(* IEC 61131-3 sources: plc-iiot-stack/adapters/sd_mqtt_1_0/src/POUs/Adapters/FB_MqttClientSdMqtt, 14 files *)

(* ---- FB_MqttClientSdMqtt.decl.st ---- *)
// Назначение: адаптер I_MqttClient на библиотеку CODESYS-MQTT (github.com/stefandreyer/CODESYS-MQTT), релиз
//             «stable» (Project Information: MQTT 1.0.0.0, компания Stefan Dreyer, пространство имён SD_MQTT).
//             НЕ КОМПИЛИРОВАЛСЯ С РАБОЧЕЙ БИБЛИОТЕКОЙ: на CODESYS 3.5.17.30 у библиотеки нет зависимостей
//             (OSCAT BASIC 3.3.3.0, OSCAT NETWORK 1.30, «Common Helper for development» и системные
//             библиотеки точных версий 3.5.5–3.5.13), поэтому файл лежит вне src/ (docs/MANUAL_STEPS.md, раздел 9).
//             Сигнатуры взяты из объявлений библиотеки (HANDLE_MQTT, MQTTPublish, MQTTSubscribe, MQTT_IN_OUT).
//             Пул из PUB_POOL публикаторов: библиотека требует не менять топик и текст до done и пускает
//             публикацию по фронту send. Логин и пароль брокера версия 1.0.0.0 через входы не принимает —
//             Connect с непустым sUser отклоняется (MQTT_ERR_AUTH_UNSUPPORTED), а не подключается без пароля.
//             Завещание (LWT) версия строит сама из ClientID (WillTopicBase, ClientWillTopic, ClientWillMessage
//             до 30 символов): offline/lwt по data_schema 6 с ней не получить; флаг retain принятых сообщений
//             не виден (проверка retained шлюза команд не срабатывает).
// Автор:      kr0nsch
// Версия:     0.1.0
// Документ:   docs/plc_mqtt.md, раздел «Адаптер I_MqttClient»
FUNCTION_BLOCK FB_MqttClientSdMqtt IMPLEMENTS I_MqttClient
VAR_INPUT
    tTimeout : TIME := T#5S;                           // HANDLE_MQTT.TIMEOUT
END_VAR
VAR
    fbHandler : SD_MQTT.HANDLE_MQTT;
    stInOut : SD_MQTT.MQTT_IN_OUT;
    stInfo : SD_MQTT.MQTT_INFO;
    aPublishers : ARRAY[1..PUB_POOL] OF SD_MQTT.MQTTPublish;
    aPubTopic : ARRAY[1..PUB_POOL] OF STRING(GVL_Const.MQTT_TOPIC_LEN);
    aPubPayload : ARRAY[1..PUB_POOL] OF STRING(GVL_Const.MQTT_PAYLOAD_LEN);
    aPubLen : ARRAY[1..PUB_POOL] OF UDINT;
    aPubQos : ARRAY[1..PUB_POOL] OF SD_MQTT.QoS;
    aPubRetain : ARRAY[1..PUB_POOL] OF BOOL;
    aPubState : ARRAY[1..PUB_POOL] OF USINT;          // SLOT_FREE, SLOT_SENDING, SLOT_RELEASE
    fbSubscriber : SD_MQTT.MQTTSubscribe;
    sSubFilter : STRING(GVL_Const.MQTT_TOPIC_LEN);
    eSubQos : SD_MQTT.QoS;
    xSubscribe : BOOL;
    aRxTopic : ARRAY[1..RX_MAX] OF STRING(GVL_Const.MQTT_TOPIC_LEN);
    aRxPayload : ARRAY[1..RX_MAX] OF STRING(GVL_Const.MQTT_CMD_PAYLOAD_LEN);
    aRxTruncated : ARRAY[1..RX_MAX] OF BOOL;
    uiRxCount : UINT;
    sUrl : STRING(GVL_Const.MQTT_TOPIC_LEN);
    xEnable : BOOL;
    xTls : BOOL;
    xBound : BOOL;                                     // SetMqttInOut выполнен у всех ФБ библиотеки
    diError : DINT;
    uiSlot : UINT;
END_VAR
VAR CONSTANT
    PUB_POOL : UINT := 8;
    RX_MAX : UINT := 8;
    SLOT_FREE : USINT := 0;
    SLOT_SENDING : USINT := 1;     // send = TRUE до done или SendTimeout
    SLOT_RELEASE : USINT := 2;     // один вызов с send = FALSE, чтобы следующий фронт был виден
    MQTT_ERR_AUTH_UNSUPPORTED : DINT := -10;
    MQTT_ERR_SEND_TIMEOUT : DINT := -11;
END_VAR

(* ---- Connect.method.decl.st ---- *)
// Адрес host:port, идентификатор клиента, TLS; логин и пароль не поддерживаются (см. заголовок).
METHOD Connect : BOOL
VAR_IN_OUT CONSTANT
    // lint:allow STL007 параметр VAR_IN_OUT CONSTANT — ссылка только для чтения, а не константа
    stCfg : ST_MqttBrokerCfg;
END_VAR

(* ---- Connect.method.impl.st ---- *)
IF LEN(stCfg.sUser) > 0 OR LEN(stCfg.sPassword) > 0 THEN
    diError := MQTT_ERR_AUTH_UNSUPPORTED;
    RETURN;
END_IF
sUrl := CONCAT(CONCAT(stCfg.sHost, ':'), UINT_TO_STRING(stCfg.uiPort));
stInOut.ClientID := stCfg.sClientId;
xTls := stCfg.xTls;
diError := GVL_Const.MQTT_ERR_NONE;
xEnable := TRUE;
Connect := TRUE;

(* ---- Cycle.method.decl.st ---- *)
// Обработчик библиотеки, публикаторы и подписчик — один раз за цикл задачи.
METHOD Cycle
VAR
    pSrc : POINTER TO BYTE;
    udiLen : UDINT;
    uiIdx : UINT;
END_VAR

(* ---- Cycle.method.impl.st ---- *)
IF NOT xBound THEN
    FOR uiSlot := 1 TO PUB_POOL DO
        aPublishers[uiSlot].SetMqttInOut(MQTT_IN_OUT := ADR(stInOut));
    END_FOR
    fbSubscriber.SetMqttInOut(MQTT_IN_OUT := ADR(stInOut));
    xBound := TRUE;
END_IF

fbHandler(ENABLE := xEnable, URL := sUrl, TIMEOUT := tTimeout, TLS := xTls, MQTT_INFO := stInfo,
    MQTT_IN_OUT := stInOut);
IF fbHandler.ERROR_C <> 0 THEN
    diError := DWORD_TO_DINT(fbHandler.ERROR_C);
END_IF

FOR uiSlot := 1 TO PUB_POOL DO
    aPublishers[uiSlot](Topic := ADR(aPubTopic[uiSlot]), PayloadString := 0, PublishAsString := FALSE,
                        Payload := ADR(aPubPayload[uiSlot]), PayloadLength := aPubLen[uiSlot], QoSIn := aPubQos[uiSlot],
                        MRetain := aPubRetain[uiSlot], send := aPubState[uiSlot] = SLOT_SENDING);
    IF aPubState[uiSlot] = SLOT_SENDING THEN
        IF aPublishers[uiSlot].SendTimeout THEN
            diError := MQTT_ERR_SEND_TIMEOUT;
            aPubState[uiSlot] := SLOT_RELEASE;
        ELSIF aPublishers[uiSlot].done THEN
            aPubState[uiSlot] := SLOT_RELEASE;
        END_IF
    ELSIF aPubState[uiSlot] = SLOT_RELEASE THEN
        aPubState[uiSlot] := SLOT_FREE;
    END_IF
END_FOR

fbSubscriber(Subscribe := xSubscribe AND IsConnected(), Topic := ADR(sSubFilter), QoSSubscribe := eSubQos,
             ExpectingString := FALSE);
IF fbSubscriber.Recived AND uiRxCount < RX_MAX AND fbSubscriber.TopicOut <> 0 AND fbSubscriber.Payload <> 0 THEN
    uiRxCount := uiRxCount + 1;
    aRxTopic[uiRxCount] := fbSubscriber.TopicOut^;
    udiLen := fbSubscriber.PayloadSize;
    aRxTruncated[uiRxCount] := udiLen > GVL_Const.MQTT_CMD_PAYLOAD_LEN;
    IF udiLen > GVL_Const.MQTT_CMD_PAYLOAD_LEN THEN
        udiLen := GVL_Const.MQTT_CMD_PAYLOAD_LEN;
    END_IF
    pSrc := fbSubscriber.Payload;
    uiIdx := 0;
    WHILE uiIdx < UDINT_TO_UINT(udiLen) DO
        aRxPayload[uiRxCount][uiIdx] := (pSrc + uiIdx)^;
        uiIdx := uiIdx + 1;
    END_WHILE
    aRxPayload[uiRxCount][uiIdx] := 0;
END_IF

(* ---- Disconnect.method.impl.st ---- *)
xEnable := FALSE;
xSubscribe := FALSE;
uiRxCount := 0;
FOR uiSlot := 1 TO PUB_POOL DO
    aPubState[uiSlot] := SLOT_FREE;
END_FOR
Disconnect := TRUE;

(* ---- Publish.method.decl.st ---- *)
// Занять свободный публикатор пула: копия топика и текста (библиотека читает их до done).
METHOD Publish : BOOL
VAR_INPUT
    sTopic : STRING(GVL_Const.MQTT_TOPIC_LEN);
    eQos : E_MqttQos;
    xRetain : BOOL;
END_VAR
VAR_IN_OUT CONSTANT
    // lint:allow STL007 параметр VAR_IN_OUT CONSTANT — ссылка только для чтения, а не константа
    sPayload : STRING(GVL_Const.MQTT_PAYLOAD_LEN);
END_VAR
VAR
    uiLen : UINT;
END_VAR

(* ---- Publish.method.impl.st ---- *)
IF NOT IsConnected() THEN
    RETURN;
END_IF
FOR uiSlot := 1 TO PUB_POOL DO
    IF aPubState[uiSlot] = SLOT_FREE THEN
        uiLen := 0;
        WHILE uiLen < GVL_Const.MQTT_PAYLOAD_LEN AND_THEN sPayload[uiLen] <> 0 DO
            uiLen := uiLen + 1;
        END_WHILE
        aPubTopic[uiSlot] := sTopic;
        aPubPayload[uiSlot] := sPayload;
        aPubLen[uiSlot] := UINT_TO_UDINT(uiLen);
        aPubQos[uiSlot] := ToLibQos(eQosIn := eQos);
        aPubRetain[uiSlot] := xRetain;
        aPubState[uiSlot] := SLOT_SENDING;
        Publish := TRUE;
        RETURN;
    END_IF
END_FOR

(* ---- Receive.method.decl.st ---- *)
// Первое принятое сообщение из очереди адаптера.
METHOD Receive : BOOL
VAR_IN_OUT
    sTopic : STRING(GVL_Const.MQTT_TOPIC_LEN);
    sPayload : STRING(GVL_Const.MQTT_CMD_PAYLOAD_LEN);
END_VAR
VAR_OUTPUT
    xTruncated : BOOL;
    xRetained : BOOL;      // версия 1.0.0.0 флаг retain принятого сообщения не отдаёт: всегда FALSE
END_VAR
VAR
    uiIdx : UINT;
END_VAR

(* ---- Receive.method.impl.st ---- *)
xRetained := FALSE;
IF uiRxCount = 0 THEN
    RETURN;
END_IF
sTopic := aRxTopic[1];
sPayload := aRxPayload[1];
xTruncated := aRxTruncated[1];
FOR uiIdx := 1 TO uiRxCount - 1 DO
    aRxTopic[uiIdx] := aRxTopic[uiIdx + 1];
    aRxPayload[uiIdx] := aRxPayload[uiIdx + 1];
    aRxTruncated[uiIdx] := aRxTruncated[uiIdx + 1];
END_FOR
uiRxCount := uiRxCount - 1;
Receive := TRUE;

(* ---- Subscribe.method.decl.st ---- *)
// Подписка одним подписчиком библиотеки (адаптеру нужен один фильтр: <prefix>/+/+/cmd).
METHOD Subscribe : BOOL
VAR_INPUT
    sTopicFilter : STRING(GVL_Const.MQTT_TOPIC_LEN);
    eQos : E_MqttQos;
END_VAR

(* ---- Subscribe.method.impl.st ---- *)
IF NOT IsConnected() THEN
    RETURN;
END_IF
sSubFilter := sTopicFilter;
eSubQos := ToLibQos(eQosIn := eQos);
xSubscribe := TRUE;
Subscribe := NOT fbSubscriber.SubscribeFail;

(* ---- ToLibQos.method.decl.st ---- *)
// E_MqttQos -> SD_MQTT.QoS.
METHOD PRIVATE ToLibQos : SD_MQTT.QoS
VAR_INPUT
    eQosIn : E_MqttQos;
END_VAR

(* ---- ToLibQos.method.impl.st ---- *)
CASE eQosIn OF
    E_MqttQos.AtLeastOnce:
        ToLibQos := SD_MQTT.QoS.AtLeastOnce;
    E_MqttQos.ExactlyOnce:
        ToLibQos := SD_MQTT.QoS.ExactlyOnce;
ELSE
    ToLibQos := SD_MQTT.QoS.AtMostOnce;
END_CASE
